Fanuc KAREL source: KT00867.KL

PROGRAM KT00867
%NOLOCKGROUP
VAR
  S1: STRING[80]
  S2: STRING[80]
  OUT: REAL
BEGIN
  S1 = 'A'
  S2 = 'B'
  S1 = 'A'
  S2 = 'B'
  OUT = ROUND(S1)
END KT00867
